FUNCTION F_RangeOpen : ST_Range		// 제한 없는 범위
VAR
END_VAR

F_RangeOpen.fMax := 1.0E30;
F_RangeOpen.fMin := -1.0E30;

END_FUNCTION

(* stored: Version 1.1.0.1, ProductVersion 3.1.4024.15
   POU F_RangeOpen: Id {f29ef760-35fa-432f-b15c-e56fb3b6e0f8}, SpecialFunc None *)
